    rq_activate_all_grippers(True)
    # end: URCap Program Node
  end
  $ 58 "zero_ftsensor()"
  zero_ftsensor()
  $ 59 "EXTT"
  $ 60 "Set GRP_3F_Enable=Off"
  set_standard_digital_out(4, False)
  $ 61 "Set BarcodeTrigger=Off"
  set_standard_digital_out(6, False)
  $ 62 "Set GRP_3F_Decap=Off"
  set_standard_digital_out(3, False)
  $ 63 "Set GRP_3F_Cap=Off"
  set_standard_digital_out(2, False)
  $ 64 "Set GRP_3F_Open=Off"
  set_standard_digital_out(5, False)
  $ 65 "PSE_T≔get_tool_free_pose(dir=[0,0,0.150], move_in_base_frame=True)"
  global PSE_T=get_tool_free_pose(dir=[0,0,0.150], move_in_base_frame=True)
  $ 66 "If is_reachable(Base_const, [PSE_T])"
  if (is_reachable(p[0.0,0.0,0.0,0.0,0.0,0.0], [PSE_T])):
    $ 67 "MoveL"
    $ 68 "PSE_T" "breakAfter"
    movel(PSE_T, a=1.2, v=0.15)
  end
  $ 69 "powder dispensing variable init"
  $ 70 "Start_thread≔ False "
  global Start_thread=  False
  $ 71 "vib_thread≔ False "
  global vib_thread=  False
  $ 72 "w_full_thread≔ False "
  global w_full_thread=  False
  $ 73 "Picking≔ False "
  global Picking=  False
  $ 74 "d_cc≔0.07"
  global d_cc=0.07
  $ 75 "kp≔0.0035"
  global kp=0.0035
  $ 76 "ki≔0.0001"
  global ki=0.0001
  $ 77 "kd≔0.003"
  global kd=0.003
  $ 78 "dt≔0.2"
  global dt=0.2
  $ 79 "Integral_error≔0"
  global Integral_error=0
  $ 80 "current_error≔0"
  global current_error=0
  $ 81 "previous_error≔0"
  global previous_error=0
  $ 82 "tilt_increment≔0"
  global tilt_increment=0
  $ 83 "tilt_angle≔0"
  global tilt_angle=0
  $ 84 "diff≔0"
  global diff=0
  $ 85 "tilt_to_home()"
  tilt_to_home()
  $ 86 "params_init()"
  params_init()
  $ 87 "switch_spat_M≔ True "
  global switch_spat_M=  True
  $ 88 "switch_spat_S≔ True "
  global switch_spat_S=  True
  $ 89 "switch_spat_F_M≔ True "
  global switch_spat_F_M=  True
  $ 90 "switch_spat_F_S≔ True "
  global switch_spat_F_S=  True
  $ 861 "Thread_1"
  thread Thread_1():
    while (True):
      $ 862 "Dosing Weight"
      $ 863 "If Start_thread≟ True "
      if (Start_thread ==   True  ):
        $ 864 "weight_value≔get_weight()"
        global weight_value=get_weight()
        $ 865 "diff≔target_weight-weight_value"
        global diff=target_weight-weight_value
        $ 866 "Wait: 0.2"
        sleep(0.2)
        $ 867 "sync()"
        sync()
      end
      $ 868 "sync()"
      sync()
    end
  end
  threadId_Thread_1 = run Thread_1()
  $ 869 "Thread_2"
  thread Thread_2():
    while (True):
      $ 883 "Vibration motor"
      $ 884 "Loop vib_thread≟ True "
      thread Thread_while_884():
        while (True):
          $ 885 "If spatula≟'spatula_S' "
          global thread_flag_885=0
          thread Thread_if_885():
            $ 886 "vibration_4()"
            vibration_4()
            thread_flag_885 = 1
          end
          if (spatula == "spatula_S" ):
            global thread_handler_885=run Thread_if_885()
            while (thread_flag_885 == 0):
              if not(spatula == "spatula_S" ):
                kill thread_handler_885
                thread_flag_885 = 2
              else:
                sync()
              end
            end
          else:
            thread_flag_885 = 2
          end
          if (thread_flag_885 == 2):
            $ 887 "ElseIf spatula≟'spatula_M'"
            if (spatula == "spatula_M"):
              $ 888 "vibration_3()"
              vibration_3()
            else:
              $ 889 "Else" "noBreak"
              $ 890 "Set AO[0]=0.0"
              set_standard_analog_out(0, 0.0)
              $ 891 "textmsg('stopped')"
              textmsg("stopped")
            end
          end
        end
      end
      if (vib_thread ==   True  ):
        global thread_handler_884=run Thread_while_884()
        while (vib_thread ==   True  ):
          sync()
        end
        kill thread_handler_884
      end
      $ 892 "sync()"
      sync()
    end
  end
  threadId_Thread_2 = run Thread_2()
  $ 893 "Thread_3"
  thread Thread_3():
    while (True):
      $ 894 "Container weight"
      $ 895 "If w_full_thread≟ True "
      if (w_full_thread ==   True  ):
        $ 896 "aa_weight_cont≔get_cont_weight()"
        global aa_weight_cont=get_cont_weight()
        $ 897 "Wait: 0.2"
        sleep(0.2)
        $ 898 "sync()"
        sync()
      end
      $ 899 "sync()"
      sync()
    end
  end
  threadId_Thread_3 = run Thread_3()
  while (True):
    $ 92 "Robot Program"
    $ 93 "MAIN"
    $ 94 "command_manager(external_control='uGO', cond_suspend=(ITM_Manipulated and AMR_AtTarget and AMR_Charging and AMR_Battery<40), cond_unsuspend=(AMR_Battery≟60))"
    command_manager(external_control="uGO", cond_suspend=(ITM_Manipulated  and  AMR_AtTarget  and  AMR_Charging  and  AMR_Battery<40), cond_unsuspend=(AMR_Battery == 60))
    $ 95 "log_state(STATE_Info)"
    log_state(STATE_Info)
    $ 96 "Switch STATE"
    switch_1 = STATE
    $ 97 "Case 1"
    if (1 == switch_1):
      $ 98 "Stopping"
      $ 99 "STATE_Info≔'Stopping'"
      global STATE_Info="Stopping"
      $ 100 "end_freedrive_mode()"
      end_freedrive_mode()
      $ 101 "Set"
      set_tcp(p[0.0,0.0,0.161,3.1415,0.0,0.0])
      $ 102 "PSE_T≔get_tool_free_pose(dir=[0,0,0.150], move_in_base_frame=True)"
      global PSE_T=get_tool_free_pose(dir=[0,0,0.150], move_in_base_frame=True)
      $ 103 "If is_reachable(Base_const, [PSE_T])"
      if (is_reachable(p[0.0,0.0,0.0,0.0,0.0,0.0], [PSE_T])):
        $ 104 "MoveL"
        $ 105 "PSE_T" "breakAfter"
        movel(PSE_T, a=1.2, v=0.15)
      end
      $ 106 "do_transition(keep_rxry=OBJ_Picked, r=0)"
      do_transition(keep_rxry=OBJ_Picked, r=0)
      $ 115 "Call Sub_AMR_MiR_V3"
      Sub_AMR_MiR_V3()
      $ 116 "If stopping() and AMR_Done"
      if (stopping()  and  AMR_Done):
        $ 117 "STATE≔2"
        global STATE=2
        $ 118 "ugo_update_outputs()"
        ugo_update_outputs()
      end
    elif (2 == switch_1):
      $ 119 "Case 2"
      $ 120 "Stopped"
      $ 121 "STATE_Info≔'Stopped'"
      global STATE_Info="Stopped"
      $ 122 "Call Sub_AMR_MiR_V3"
      Sub_AMR_MiR_V3()
      $ 123 "If CMD_Reset  or PB_Start"
      if (CMD_Reset   or  get_standard_digital_in(0)):
        $ 124 "STATE≔3"
        global STATE=3
        $ 125 "ugo_update_outputs()"
        ugo_update_outputs()
      end
    elif (3 == switch_1):
      $ 126 "Case 3"
      $ 127 " Resetting"
      $ 128 "STATE_Info≔'Resetting'"
      global STATE_Info="Resetting"
      $ 129 "uML"
      $ 130 "reset_error()"
      reset_error()
      $ 131 "reset_warning()"
      reset_warning()
      $ 132 "PROCESS_Step≔0"
      global PROCESS_Step=0
      $ 133 "PROCESS_Info≔''"
      global PROCESS_Info=""
      $ 134 "ARM_Referenced≔ False "
      global ARM_Referenced=  False
      $ 135 "WRK_Done≔ False "
      global WRK_Done=  False
      $ 136 "ITM_Prepared≔ False "
      global ITM_Prepared=  False
      $ 137 "ITM_Manipulated≔ False "
      global ITM_Manipulated=  False
      $ 138 "STP≔0"
      global STP=0
      $ 139 "Action≔0"
      global Action=0
      $ 140 "Action_Info≔''"
      global Action_Info=""
      $ 141 "ITM_ID≔0"
      global ITM_ID=0
      $ 142 "JIG≔0"
      global JIG=0
      $ 143 "JIG_Slot≔0"
      global JIG_Slot=0
      $ 144 "Task_info≔''"
      global Task_info=""
      $ 145 "Set"
      set_tcp(p[0.0,0.0,0.161,3.1415,0.0,0.0])
      $ 146 "App"
      $ 147 "'ADD APPLICATION SPECIFIC COMMANDS'"
      # 'ADD APPLICATION SPECIFIC COMMANDS'
      $ 148 "OBJ_Type≔0"
      global OBJ_Type=0
      $ 149 "OBJ_Nbr≔0"
      global OBJ_Nbr=0
      $ 150 "If CNT_Rack_Output≥50"
      if (CNT_Rack_Output >= 50):
        $ 151 "CNT_Rack_Output≔0"
        global CNT_Rack_Output=0
      end
      $ 152 "TASK≔struct(ID=0, NAVI=struct(target=0, footprint=0, protectiveOff=0, dock=0), WORK=struct(ITM_ID_Src=0, JIG_ID_Src=0, OBJ_Nbr_Src=0, ACT_Src=0, ITM_ID_Tgt=0, JIG_ID_Tgt=0, OBJ_Nbr_Tgt=0, ACT_Tgt=0, OBJ_Type=0))"
      global TASK=struct(ID=0, NAVI=struct(target=0, footprint=0, protectiveOff=0, dock=0), WORK=struct(ITM_ID_Src=0, JIG_ID_Src=0, OBJ_Nbr_Src=0, ACT_Src=0, ITM_ID_Tgt=0, JIG_ID_Tgt=0, OBJ_Nbr_Tgt=0, ACT_Tgt=0, OBJ_Type=0))
      $ 153 "Call Sub_AMR_MiR_V3"
      Sub_AMR_MiR_V3()
      $ 154 "If resetting() and AMR_Done"
      if (resetting()  and  AMR_Done):
        $ 155 "STATE≔4"
        global STATE=4
        $ 156 "ugo_update_outputs()"
        ugo_update_outputs()
      end
    elif (4 == switch_1):
      $ 157 "Case 4"
      $ 158 "Idle"
      $ 159 "STATE_Info≔'Idle'"
      global STATE_Info="Idle"
      $ 160 "If CMD_Start"
      if (CMD_Start):
        $ 161 "STATE≔5"
        global STATE=5
        $ 162 "ugo_update_outputs()"
        ugo_update_outputs()
      end
    elif (5 == switch_1):
      $ 163 "Case 5"
      $ 164 "Starting"
      $ 165 "STATE_Info≔'Starting'"
      global STATE_Info="Starting"
      $ 166 "'ADD COMMANDS WHAT TO START WITH'"
      # 'ADD COMMANDS WHAT TO START WITH'
      $ 167 "Call Sub_AMR_MiR_V3"
      Sub_AMR_MiR_V3()
      $ 168 "get ugo data"
      $ 169 "Assign Tasks"
      $ 170 "TASK.ID = ugo_get_task()"
      TASK.ID = ugo_get_task()
      $ 171 "If TASK.ID≟1"
      if (TASK.ID == 1):
        $ 172 "Task_info≔'Charge'"
        global Task_info="Charge"
        $ 173 "Parameters"
        $ 174 "AMR_PosTarget≔1"
        global AMR_PosTarget=1
      else:
        $ 175 "ElseIf TASK.ID≟9"
        if (TASK.ID == 9):
          $ 176 "'Pick Sarstedt Rack from Variable source'"
          # 'Pick Sarstedt Rack from Variable source'
          $ 177 "Task_info≔'Navigate to Target'"
          global Task_info="Navigate to Target"
          $ 178 "Parameters"
          $ 179 "AMR_PosTarget≔UGO.read_input('00','ITM_ID')"
          global AMR_PosTarget=UGO.read_input("00","ITM_ID")
        else:
          $ 180 "ElseIf TASK.ID≟13"
          if (TASK.ID == 13):
            $ 181 "Task_info≔'Dose Powder'"
            global Task_info="Dose Powder"
            $ 182 "Parameters"
            $ 183 "ITM_ID≔1"
            global ITM_ID=1
            $ 184 "W_now≔(UGO.read_input('00','Container_weight'))/1000"
            global W_now=(UGO.read_input("00","Container_weight"))/1000
            $ 185 "Pow_name≔(UGO.read_input('00','Powder_name'))"
            global Pow_name=(UGO.read_input("00","Powder_name"))
            $ 186 "target_weight≔(UGO.read_input('00','Target_weight'))/1000"
            global target_weight=(UGO.read_input("00","Target_weight"))/1000
            $ 187 "params_init()"
            params_init()
            $ 188 "send_picking_info(Pow_name,target_weight)"
            send_picking_info(Pow_name,target_weight)
            $ 190 "OBJ_Type≔6"
            global OBJ_Type=6
            $ 191 "JIG≔17"
            global JIG=17
            $ 192 "AMR_PosTarget≔5"
            global AMR_PosTarget=5
          else:
            $ 193 "ElseIf TASK.ID≟49"
            if (TASK.ID == 49):
              $ 194 "Task_info≔'Pick Containers'"
              global Task_info="Pick Containers"
              $ 195 "Parameters"
              $ 196 "ITM_ID≔1"
              global ITM_ID=1
              $ 197 "OBJ_Type≔6"
              global OBJ_Type=6
              $ 198 "JIG≔15"
              global JIG=15
              $ 199 "AMR_PosTarget≔3"
              global AMR_PosTarget=3
            else:
              $ 200 "ElseIf TASK.ID≟50"
              if (TASK.ID == 50):
                $ 201 "Task_info≔'Decap Containers'"
                global Task_info="Decap Containers"
                $ 202 "Parameters"
                $ 203 "ITM_ID≔1"
                global ITM_ID=1
                $ 204 "OBJ_Type≔6"
                global OBJ_Type=6
                $ 205 "JIG≔16"
                global JIG=16
                $ 206 "AMR_PosTarget≔5"
                global AMR_PosTarget=5
              else:
                $ 207 "ElseIf TASK.ID≟51"
                if (TASK.ID == 51):
                  $ 208 "Task_info≔'Detect Spatula and transfer powder'"
                  global Task_info="Detect Spatula and transfer powder"
                  $ 209 "Parameters"
                  $ 210 "ITM_ID≔1"
                  global ITM_ID=1
                  $ 211 "target_weight≔(UGO.read_input('00','Target_weight'))/1000"
                  global target_weight=(UGO.read_input("00","Target_weight"))/1000
                  $ 212 "OBJ_Type≔8"
                  global OBJ_Type=8
                  $ 213 "JIG≔16"
                  global JIG=16
                  $ 214 "AMR_PosTarget≔5"
                  global AMR_PosTarget=5
                else:
                  $ 215 "ElseIf TASK.ID≟52"
                  if (TASK.ID == 52):
                    $ 216 "Task_info≔'Pick Powder'"
                    global Task_info="Pick Powder"
                    $ 217 "Parameters"
                    $ 218 "ITM_ID≔1"
                    global ITM_ID=1
                    $ 220 "OBJ_Type≔6"
                    global OBJ_Type=6
                    $ 221 "JIG≔15"
                    global JIG=15
                    $ 222 "AMR_PosTarget≔3"
                    global AMR_PosTarget=3
                  else:
                    $ 223 "ElseIf TASK.ID≟53"
                    if (TASK.ID == 53):
                      $ 224 "Task_info≔'Decap Powder'"
                      global Task_info="Decap Powder"
                      $ 225 "Parameters"
                      $ 226 "ITM_ID≔1"
                      global ITM_ID=1
                      $ 227 "OBJ_Type≔6"
                      global OBJ_Type=6
                      $ 228 "JIG≔1"
                      global JIG=1
                      $ 229 "AMR_PosTarget≔5"
                      global AMR_PosTarget=5
                    else:
                      $ 230 "ElseIf TASK.ID≟54"
                      if (TASK.ID == 54):
                        $ 231 "Task_info≔'Empty and swap Powder container'"
                        global Task_info="Empty and swap Powder container"
                        $ 240 "Parameters"
                        $ 241 "ITM_ID≔1"
                        global ITM_ID=1
                        $ 243 "W_now≔(UGO.read_input('00','Container_weight'))/1000"
                        global W_now=(UGO.read_input("00","Container_weight"))/1000
                        $ 244 "Pow_name≔(UGO.read_input('00','Powder_name'))"
                        global Pow_name=(UGO.read_input("00","Powder_name"))
                        $ 247 "OBJ_Type≔6"
                        global OBJ_Type=6
                        $ 248 "JIG≔17"
                        global JIG=17
                        $ 249 "AMR_PosTarget≔5"
                        global AMR_PosTarget=5
                      else:
                        $ 250 "ElseIf TASK.ID≟55"
                        if (TASK.ID == 55):
                          $ 251 "Task_info≔'Place Powder'"
                          global Task_info="Place Powder"
                          $ 252 "Parameters"
                          $ 253 "ITM_ID≔1"
                          global ITM_ID=1
                          $ 254 "OBJ_Type≔6"
                          global OBJ_Type=6
                          $ 255 "JIG≔21"
                          global JIG=21
                          $ 256 "AMR_PosTarget≔5"
                          global AMR_PosTarget=5
                        else:
                          $ 257 "ElseIf TASK.ID≟56"
                          if (TASK.ID == 56):
                            $ 258 "Task_info≔'Dose Powder'"
                            global Task_info="Dose Powder"
                            $ 259 "Parameters"
                            $ 260 "ITM_ID≔1"
                            global ITM_ID=1
                            $ 261 "target_weight≔(UGO.read_input('00','Target_weight'))/1000"
                            global target_weight=(UGO.read_input("00","Target_weight"))/1000
                            $ 262 "W_now≔(UGO.read_input('00','Container_weight'))/1000"
                            global W_now=(UGO.read_input("00","Container_weight"))/1000
                            $ 263 "Pow_name≔(UGO.read_input('00','Powder_name'))"
                            global Pow_name=(UGO.read_input("00","Powder_name"))
                            $ 264 "OBJ_Type≔6"
                            global OBJ_Type=6
                            $ 265 "JIG≔17"
                            global JIG=17
                            $ 266 "AMR_PosTarget≔5"
                            global AMR_PosTarget=5
                          else:
                            $ 267 "ElseIf TASK.ID≟57"
                            if (TASK.ID == 57):
                              $ 268 "Task_info≔'Recipe Powder dosing'"
                              global Task_info="Recipe Powder dosing"
                              $ 269 "Parameters"
                              $ 270 "ITM_ID≔1"
                              global ITM_ID=1
                              $ 271 "Pow_A≔(UGO.read_input('00','PowderA'))"
                              global Pow_A=(UGO.read_input("00","PowderA"))
                              $ 272 "Pow_B≔(UGO.read_input('00','PowderB'))"
                              global Pow_B=(UGO.read_input("00","PowderB"))
                              $ 273 "Pow_C≔(UGO.read_input('00','PowderC'))"
                              global Pow_C=(UGO.read_input("00","PowderC"))
                              $ 274 "Total_weight≔(UGO.read_input('00','Total_weight'))/1000"
                              global Total_weight=(UGO.read_input("00","Total_weight"))/1000
                              $ 275 "Pow_A_percent≔(UGO.read_input('00','PowderA_percentage'))/100"
                              global Pow_A_percent=(UGO.read_input("00","PowderA_percentage"))/100
                              $ 276 "Pow_B_percent≔(UGO.read_input('00','PowderB_percentage'))/100"
                              global Pow_B_percent=(UGO.read_input("00","PowderB_percentage"))/100
                              $ 277 "Pow_C_percent≔(UGO.read_input('00','PowderC_percentage'))/100"
                              global Pow_C_percent=(UGO.read_input("00","PowderC_percentage"))/100
                              $ 278 "OBJ_Type≔6"
                              global OBJ_Type=6
                              $ 279 "JIG≔17"
                              global JIG=17
                              $ 280 "AMR_PosTarget≔5"
                              global AMR_PosTarget=5
                            else:
                              $ 281 "ElseIf TASK.ID≟58"
                              if (TASK.ID == 58):
                                $ 282 "Task_info≔'Pick Powder containers'"
                                global Task_info="Pick Powder containers"
                                $ 283 "Parameters"
                                $ 284 "ITM_ID≔1"
                                global ITM_ID=1
                                $ 285 "OBJ_Type≔6"
                                global OBJ_Type=6
                                $ 286 "JIG≔15"
                                global JIG=15
                                $ 287 "AMR_PosTarget≔3"
                                global AMR_PosTarget=3
                              else:
                                $ 288 "ElseIf TASK.ID≟59"
                                if (TASK.ID == 59):
                                  $ 289 "Task_info≔'Empty Powder container'"
                                  global Task_info="Empty Powder container"
                                  $ 290 "Parameters"
                                  $ 291 "ITM_ID≔1"
                                  global ITM_ID=1
                                  $ 293 "Pow_name≔(UGO.read_input('00','Powder_name'))"
                                  global Pow_name=(UGO.read_input("00","Powder_name"))
                                  $ 295 "target_weight≔(aa_weight_cont-empty_weight_g)"
                                  global target_weight=(aa_weight_cont-empty_weight_g)
                                  $ 296 "W_now≔target_weight"
                                  global W_now=target_weight
                                  $ 297 "params_init()"
                                  params_init()
                                  $ 298 "send_picking_info(Pow_name,target_weight)"
                                  send_picking_info(Pow_name,target_weight)
                                  $ 299 "w_dosed_total≔0"
                                  global w_dosed_total=0
                                  $ 300 "OBJ_Type≔6"
                                  global OBJ_Type=6
                                  $ 301 "JIG≔17"
                                  global JIG=17
                                  $ 302 "AMR_PosTarget≔5"
                                  global AMR_PosTarget=5
                                else:
                                  $ 303 "ElseIf TASK.ID≟61"
                                  if (TASK.ID == 61):
                                    $ 304 "Task_info≔'Weigh, Place & Decap'"
                                    global Task_info="Weigh, Place & Decap"
                                    $ 305 "Parameters"
                                    $ 306 "ITM_ID≔1"
                                    global ITM_ID=1
                                    $ 307 "OBJ_Type≔6"
                                    global OBJ_Type=6
                                    $ 308 "JIG≔21"
                                    global JIG=21
                                    $ 309 "AMR_PosTarget≔5"
                                    global AMR_PosTarget=5
                                  else:
                                    $ 310 "ElseIf TASK.ID≟62"
                                    if (TASK.ID == 62):
                                      $ 311 "Task_info≔'Dose Powder'"
                                      global Task_info="Dose Powder"
                                      $ 312 "Parameters"
                                      $ 313 "ITM_ID≔1"
                                      global ITM_ID=1
                                      $ 315 "W_now≔aa_weight_cont"
                                      global W_now=aa_weight_cont
                                      $ 316 "Pow_name≔(UGO.read_input('00','Powder_name'))"
                                      global Pow_name=(UGO.read_input("00","Powder_name"))
                                      $ 317 "target_weight≔(UGO.read_input('00','Target_weight'))/1000"
                                      global target_weight=(UGO.read_input("00","Target_weight"))/1000
                                      $ 319 "params_init()"
                                      params_init()
                                      $ 320 "send_picking_info(Pow_name,target_weight)"
                                      send_picking_info(Pow_name,target_weight)
                                      $ 321 "OBJ_Type≔6"
                                      global OBJ_Type=6
                                      $ 322 "JIG≔17"
                                      global JIG=17
                                      $ 323 "AMR_PosTarget≔5"
                                      global AMR_PosTarget=5
                                    else:
                                      $ 324 "ElseIf TASK.ID≟64"
                                      if (TASK.ID == 64):
                                        $ 325 "Task_info≔'Dosing Fumehood'"
                                        global Task_info="Dosing Fumehood"
                                        $ 326 "Parameters"
                                        $ 327 "ITM_ID≔1"
                                        global ITM_ID=1
                                        $ 328 "W_now≔(UGO.read_input('00','Container_weight'))/1000"
                                        global W_now=(UGO.read_input("00","Container_weight"))/1000
                                        $ 329 "OBJ_Type≔6"
                                        global OBJ_Type=6
                                        $ 330 "JIG≔21"
                                        global JIG=21
                                        $ 331 "AMR_PosTarget≔6"
                                        global AMR_PosTarget=6
                                      else:
                                        $ 332 "Else" "noBreak"
                                        $ 333 "set_error(ERROR_WRONG_ORDER)"
                                        set_error(ERROR_WRONG_ORDER)
                                      end
                                    end
                                  end
                                end
                              end
                            end
                          end
                        end
                      end
                    end
                  end
                end
              end
            end
          end
        end
      end
      $ 334 "test ugo"
      $ 335 "Wait: 0.2"
      sleep(0.2)
      $ 336 "ugo_update_outputs()"
      ugo_update_outputs()
      $ 337 "If starting() and AMR_Done"
      if (starting()  and  AMR_Done):
        $ 338 "log_message(Task_info, 'New Task: ')"
        log_message(Task_info, "New Task: ")
        $ 339 "log_message(to_str(TASK.ID), 'Task_ID: ')"
        log_message(to_str(TASK.ID), "Task_ID: ")
        $ 340 "do_transition(keep_rxry=OBJ_Picked)"
        do_transition(keep_rxry=OBJ_Picked)
        $ 341 "STATE≔6"
        global STATE=6
        $ 342 "ugo_update_outputs()"
        ugo_update_outputs()
      end
    elif (6 == switch_1):
      $ 343 "Case 6"
      $ 344 "Execute"
      $ 345 "STATE_Info≔'Execute'"
      global STATE_Info="Execute"
      $ 346 "If  not CMD_Hold and not CMD_Suspend"
      global thread_flag_346=0
      thread Thread_if_346():
        $ 347 "Switch PROCESS_Step"
        switch_2 = PROCESS_Step
        $ 348 "Case 0"
        if (0 == switch_2):
          $ 349 "PROCESS_Info≔'process control'"
          global PROCESS_Info="process control"
          $ 350 "log_process(PROCESS_Info)"
          log_process(PROCESS_Info)
          $ 351 "process control"
          $ 352 "If  not AMR_AtTarget"
          if (  not  AMR_AtTarget):
            $ 353 "PROCESS_Step≔1"
            global PROCESS_Step=1
          else:
            $ 354 "ElseIf (( not ITM_Prepared and  not WRK_Done) or (ITM_Prepared and WRK_Done))"
            if (((  not  ITM_Prepared  and    not  WRK_Done)  or  (ITM_Prepared  and  WRK_Done))):
              $ 355 "PROCESS_Step≔2"
              global PROCESS_Step=2
            else:
              $ 356 "ElseIf  not WRK_Done"
              if (  not  WRK_Done):
                $ 357 "PROCESS_Step≔3"
                global PROCESS_Step=3
              else:
                $ 358 "Else" "noBreak"
                $ 359 "task finished"
                $ 360 "PROCESS_Info≔''"
                global PROCESS_Info=""
                $ 361 "STATE≔7"
                global STATE=7
                $ 362 "ugo_update_outputs()"
                ugo_update_outputs()
              end
            end
          end
        elif (1 == switch_2):
          $ 363 "Case 1"
          $ 364 "navigate"
          $ 365 "'MOVING THE uML'"
          # 'MOVING THE uML'
          $ 366 "PROCESS_Info≔'move to target'"
          global PROCESS_Info="move to target"
          $ 367 "log_process(PROCESS_Info)"
          log_process(PROCESS_Info)
          $ 368 "If TASK.ID≟1"
          if (TASK.ID == 1):
            $ 369 "Action≔51"
            global Action=51
          else:
            $ 370 "Else" "noBreak"
            $ 371 "Action≔52"
            global Action=52
          end
          $ 372 "Call Sub_AMR_MiR_V3"
          Sub_AMR_MiR_V3()
          $ 373 "If AMR_Done"
          if (AMR_Done):
            $ 374 "PROCESS_Step≔0"
            global PROCESS_Step=0
          end
        elif (2 == switch_2):
          $ 375 "Case 2"
          $ 376 "prepare"
          $ 377 "'THINGS THAT HAVE TO BE DONE ONCE IN A SEQUENCE,WORKFLOW'"
          # 'THINGS THAT HAVE TO BE DONE ONCE IN A SEQUENCE,WORKFLOW'
          $ 378 "PROCESS_Info≔'prepare for work'"
          global PROCESS_Info="prepare for work"
          $ 379 "log_process(PROCESS_Info)"
          log_process(PROCESS_Info)
          $ 380 "If TASK.WORK.ITM_ID_Src>1"
          if (TASK.WORK.ITM_ID_Src>1):
            $ 381 "ITM_ID≔TASK.WORK.ITM_ID_Src"
            global ITM_ID=TASK.WORK.ITM_ID_Src
          else:
            $ 382 "ElseIf TASK.WORK.ITM_ID_Tgt>1"
            if (TASK.WORK.ITM_ID_Tgt>1):
              $ 383 "ITM_ID≔TASK.WORK.ITM_ID_Tgt"
              global ITM_ID=TASK.WORK.ITM_ID_Tgt
            end
          end
          $ 384 "If  not ARM_Referenced and (ITM_ID≠0)"
          if (  not  ARM_Referenced  and  (ITM_ID != 0)):
            $ 385 "STP≔1"
            global STP=1
          else:
            $ 386 "ElseIf ARM_Referenced or (ITM_ID≟0)"
            if (ARM_Referenced  or  (ITM_ID == 0)):
              $ 387 "STP≔2"
              global STP=2
            end
          end
          $ 388 "Switch STP"
          switch_3 = STP
          $ 389 "Case 1"
          if (1 == switch_3):
            $ 390 "reference"
            $ 391 "STP_Info≔'reference at target position'"
            global STP_Info="reference at target position"
            $ 392 "log_step(STP_Info)"
            log_step(STP_Info)
            $ 393 "If ITM_ID≟1"
            if (ITM_ID == 1):
              $ 394 "CAM_Done≔ True "
              global CAM_Done=  True
            else:
              $ 395 "Else" "noBreak"
              $ 396 "Action≔131"
              global Action=131
              $ 397 "Call Sub_Vision_V18"
              Sub_Vision_V18()
            end
            $ 399 "If CAM_Done and  not ERROR.FLAG"
            if (CAM_Done  and    not  ERROR.FLAG):
              $ 400 "log_step('ARM referenced')"
              log_step("ARM referenced")
              $ 401 "ARM_Referenced≔ True "
              global ARM_Referenced=  True
            end
          elif (2 == switch_3):
            $ 402 "Case 2"
            $ 403 "manipulate"
            $ 404 "STP_Info≔'manipulate item'"
            global STP_Info="manipulate item"
            $ 405 "log_step(STP_Info)"
            log_step(STP_Info)
            $ 406 "'In case pressing button is needed'"
            # 'In case pressing button is needed'
            $ 407 "If found_in_list(ITM_ID, ITM_ID_List)"
            if (found_in_list(ITM_ID, ITM_ID_List)):
              $ 408 "Switch ITM_ID"
              switch_4 = ITM_ID
              $ 409 "Case 0"
              if (0 == switch_4):
                $ 410 "ITM_Manipulated≔ not ITM_Manipulated"
                global ITM_Manipulated=  not  ITM_Manipulated
              elif (1 == switch_4):
                $ 411 "Case 1"
                $ 412 "ITM_Manipulated≔ not ITM_Manipulated"
                global ITM_Manipulated=  not  ITM_Manipulated
              elif (2 == switch_4):
                $ 413 "Case 2"
              else:
                $ 423 "Default Case"
                $ 424 "ITM_Manipulated≔ not ITM_Manipulated"
                global ITM_Manipulated=  not  ITM_Manipulated
              end
            end
          end
          $ 425 "ITM_Prepared≔(ITM_Manipulated or  not found_in_list(ITM_ID, ITM_ID_List)) and (ARM_Referenced or ITM_ID≟0) and  not WRK_Done"
          global ITM_Prepared=(ITM_Manipulated  or    not  found_in_list(ITM_ID, ITM_ID_List))  and  (ARM_Referenced  or  ITM_ID == 0)  and    not  WRK_Done
          $ 426 "STP≔0"
          global STP=0
          $ 427 "STP_Info≔''"
          global STP_Info=""
          $ 428 "PROCESS_Step≔0"
          global PROCESS_Step=0
        elif (3 == switch_2):
          $ 429 "Case 3"
          $ 430 "work"
          $ 431 "'ADD EVERY MACHINE, OBJECT, STATION TO WORK ON'"
          # 'ADD EVERY MACHINE, OBJECT, STATION TO WORK ON'
          $ 432 "Switch ITM_ID"
          switch_3 = ITM_ID
          $ 433 "Case 1"
          if (1 == switch_3):
            $ 434 "uLM"
            $ 435 "If TASK.ID≟12"
            if (TASK.ID == 12):
              $ 436 "fill racks"
              $ 437 "Action≔151"
              global Action=151
              $ 438 "Call Sub_Vision_V18"
              Sub_Vision_V18()
              $ 439 "If  not ERROR.FLAG"
              if (  not  ERROR.FLAG):
                $ 440 "Actions for the task"
                $ 441 "Action≔1"
                global Action=1
                $ 442 "JIG≔2"
                global JIG=2
                $ 443 "JIG_Slot≔CAM_Result[0]"
                global JIG_Slot=CAM_Result[0]
                $ 444 "OBJ_Nbr≔CAM_Result[0]"
                global OBJ_Nbr=CAM_Result[0]
                $ 445 "OBJ_Type≔2"
                global OBJ_Type=2
                $ 446 "Call Sub_Action_V4"
                Sub_Action_V4()
                $ 447 "If OBJ_Picked"
                if (OBJ_Picked):
                  $ 448 "CAM_Result.remove(0)"
                  CAM_Result.remove(0)
                  $ 449 "PRC_TubCounter≔PRC_TubCounter+1"
                  global PRC_TubCounter=PRC_TubCounter+1
                  $ 450 "If PRC_TubCounter%4≟0"
                  if (PRC_TubCounter%4 == 0):
                    $ 451 "JIG_Slot≔4"
                    global JIG_Slot=4
                  else:
                    $ 452 "Else" "noBreak"
                    $ 453 "JIG_Slot≔PRC_TubCounter%4"
                    global JIG_Slot=PRC_TubCounter%4
                  end
                  $ 454 "OBJ_Nbr≔ceil(PRC_TubCounter/4)"
                  global OBJ_Nbr=ceil(PRC_TubCounter/4)
                  $ 455 "Action≔2"
                  global Action=2
                  $ 456 "JIG≔4"
                  global JIG=4
                  $ 457 "Call Sub_Action_V4"
                  Sub_Action_V4()
                  $ 458 "Action≔151"
                  global Action=151
                  $ 459 "Call Sub_Vision_V18"
                  Sub_Vision_V18()
                end
              end
              $ 460 "If (CAM_Captures≥CAM_PRM_Retries) or (PRC_TubCounter≥32)"
              if ((CAM_Captures >= CAM_PRM_Retries)  or  (PRC_TubCounter >= 32)):
                $ 461 "PROCESS_Step≔0"
                global PROCESS_Step=0
                $ 462 "WRK_Done≔ True "
                global WRK_Done=  True
              end
            else:
              $ 463 "ElseIf TASK.ID≟13"
              if (TASK.ID == 13):
                $ 464 "Dose Powder"
                $ 465 "Action≔131"
                global Action=131
                $ 466 "Call Sub_Vision_V18"
                Sub_Vision_V18()
                $ 467 "Action≔34"
                global Action=34
                $ 468 "Call Sub_Action_V4"
                Sub_Action_V4()
                $ 469 "PROCESS_Step≔0"
                global PROCESS_Step=0
                $ 470 "WRK_Done≔ True "
                global WRK_Done=  True
              else:
                $ 471 "ElseIf TASK.ID≟49"
                if (TASK.ID == 49):
                  $ 472 "Pick Powder container"
                  $ 473 "Action≔131"
                  global Action=131
                  $ 474 "Call Sub_Vision_V18"
                  Sub_Vision_V18()
                  $ 475 "Action≔35"
                  global Action=35
                  $ 476 "Call Sub_Action_V4"
                  Sub_Action_V4()
                  $ 477 "PROCESS_Step≔0"
                  global PROCESS_Step=0
                  $ 478 "WRK_Done≔ True "
                  global WRK_Done=  True
                else:
                  $ 479 "ElseIf TASK.ID≟50"
                  if (TASK.ID == 50):
                    $ 480 "Decap containers"
                    $ 481 "Action≔36"
                    global Action=36
                    $ 482 "Call Sub_Action_V4"
                    Sub_Action_V4()
                    $ 483 "PROCESS_Step≔0"
                    global PROCESS_Step=0
                    $ 484 "WRK_Done≔ True "
                    global WRK_Done=  True
                  else:
                    $ 485 "ElseIf TASK.ID≟51"
                    if (TASK.ID == 51):
                      $ 486 "Detect Spatula and transfer powder"
                      $ 487 "Action≔131"
                      global Action=131
                      $ 488 "Call Sub_Vision_V18"
                      Sub_Vision_V18()
                      $ 489 "Action≔37"
                      global Action=37
                      $ 490 "Call Sub_Action_V4"
                      Sub_Action_V4()
                      $ 491 "PROCESS_Step≔0"
                      global PROCESS_Step=0
                      $ 492 "WRK_Done≔ True "
                      global WRK_Done=  True
                    else:
                      $ 493 "ElseIf TASK.ID≟52"
                      if (TASK.ID == 52):
                        $ 494 "Pick Powder container"
                        $ 495 "Action≔131"
                        global Action=131
                        $ 496 "Call Sub_Vision_V18"
                        Sub_Vision_V18()
                        $ 497 "Action≔39"
                        global Action=39
                        $ 498 "Call Sub_Action_V4"
                        Sub_Action_V4()
                        $ 499 "PROCESS_Step≔0"
                        global PROCESS_Step=0
                        $ 500 "WRK_Done≔ True "
                        global WRK_Done=  True
                      else:
                        $ 501 "ElseIf TASK.ID≟53"
                        if (TASK.ID == 53):
                          $ 502 "Decap containerA"
                          $ 503 "Action≔40"
                          global Action=40
                          $ 504 "Call Sub_Action_V4"
                          Sub_Action_V4()
                          $ 505 "PROCESS_Step≔0"
                          global PROCESS_Step=0
                          $ 506 "WRK_Done≔ True "
                          global WRK_Done=  True
                        else:
                          $ 507 "ElseIf TASK.ID≟55"
                          if (TASK.ID == 55):
                            $ 508 "Place Powder"
                            $ 509 "Action≔131"
                            global Action=131
                            $ 510 "Call Sub_Vision_V18"
                            Sub_Vision_V18()
                            $ 511 "Action≔41"
                            global Action=41
                            $ 512 "Call Sub_Action_V4"
                            Sub_Action_V4()
                            $ 513 "PROCESS_Step≔0"
                            global PROCESS_Step=0
                            $ 514 "WRK_Done≔ True "
                            global WRK_Done=  True
                          else:
                            $ 515 "ElseIf TASK.ID≟54"
                            if (TASK.ID == 54):
                              $ 516 "Empty and swap container"
                              $ 517 "Action≔131"
                              global Action=131
                              $ 518 "Call Sub_Vision_V18"
                              Sub_Vision_V18()
                              $ 519 "Action≔42"
                              global Action=42
                              $ 520 "Call Sub_Action_V4"
                              Sub_Action_V4()
                              $ 521 "PROCESS_Step≔0"
                              global PROCESS_Step=0
                              $ 522 "WRK_Done≔ True "
                              global WRK_Done=  True
                            else:
                              $ 523 "ElseIf TASK.ID≟56"
                              if (TASK.ID == 56):
                                $ 524 "Dispense Powder"
                                $ 525 "Action≔131"
                                global Action=131
                                $ 526 "Call Sub_Vision_V18"
                                Sub_Vision_V18()
                                $ 527 "Action≔43"
                                global Action=43
                                $ 528 "Call Sub_Action_V4"
                                Sub_Action_V4()
                                $ 529 "PROCESS_Step≔0"
                                global PROCESS_Step=0
                                $ 530 "WRK_Done≔ True "
                                global WRK_Done=  True
                              else:
                                $ 531 "ElseIf TASK.ID≟57"
                                if (TASK.ID == 57):
                                  $ 532 "Recipe Dosing"
                                  $ 533 "Action≔48"
                                  global Action=48
                                  $ 534 "Call Sub_Action_V4"
                                  Sub_Action_V4()
                                  $ 551 "PROCESS_Step≔0"
                                  global PROCESS_Step=0
                                  $ 552 "WRK_Done≔ True "
                                  global WRK_Done=  True
                                else:
                                  $ 553 "ElseIf TASK.ID≟58"
                                  if (TASK.ID == 58):
                                    $ 554 "Pick Powder containers"
                                    $ 555 "Num_cont_picked≔0"
                                    global Num_cont_picked=0
                                    $ 556 "powder_position≔'Position1'"
                                    global powder_position="Position1"
                                    $ 557 "Loop Num_cont_picked<3"
                                    while (Num_cont_picked<3):
                                      $ 558 "Action≔131"
                                      global Action=131
                                      $ 559 "Call Sub_Vision_V18"
                                      Sub_Vision_V18()
                                      $ 560 "Action≔47"
                                      global Action=47
                                      $ 561 "Call Sub_Action_V4"
                                      Sub_Action_V4()
                                    end
                                    $ 562 "PROCESS_Step≔0"
                                    global PROCESS_Step=0
                                    $ 563 "WRK_Done≔ True "
                                    global WRK_Done=  True
                                  else:
                                    $ 564 "ElseIf TASK.ID≟59"
                                    if (TASK.ID == 59):
                                      $ 565 "Empty powder container"
                                      $ 566 "Action≔131"
                                      global Action=131
                                      $ 567 "Call Sub_Vision_V18"
                                      Sub_Vision_V18()
                                      $ 568 "Action≔50"
                                      global Action=50
                                      $ 569 "Call Sub_Action_V4"
                                      Sub_Action_V4()
                                      $ 570 "PROCESS_Step≔0"
                                      global PROCESS_Step=0
                                      $ 571 "WRK_Done≔ True "
                                      global WRK_Done=  True
                                    else:
                                      $ 572 "ElseIf TASK.ID≟61"
                                      if (TASK.ID == 61):
                                        $ 573 "Place Powder"
                                        $ 574 "Action≔131"
                                        global Action=131
                                        $ 575 "Call Sub_Vision_V18"
                                        Sub_Vision_V18()
                                        $ 576 "Action≔51"
                                        global Action=51
                                        $ 577 "Call Sub_Action_V4"
                                        Sub_Action_V4()
                                        $ 578 "PROCESS_Step≔0"
                                        global PROCESS_Step=0
                                        $ 579 "WRK_Done≔ True "
                                        global WRK_Done=  True
                                      else:
                                        $ 580 "ElseIf TASK.ID≟62"
                                        if (TASK.ID == 62):
                                          $ 581 "Dose Powder"
                                          $ 582 "Action≔131"
                                          global Action=131
                                          $ 583 "Call Sub_Vision_V18"
                                          Sub_Vision_V18()
                                          $ 584 "Action≔52"
                                          global Action=52
                                          $ 585 "Call Sub_Action_V4"
                                          Sub_Action_V4()
                                          $ 586 "PROCESS_Step≔0"
                                          global PROCESS_Step=0
                                          $ 587 "WRK_Done≔ True "
                                          global WRK_Done=  True
                                        else:
                                          $ 588 "ElseIf TASK.ID≟64"
                                          if (TASK.ID == 64):
                                            $ 589 "Fumehood Powder dose"
                                            $ 590 "Action≔131"
                                            global Action=131
                                            $ 591 "Call Sub_Vision_V18"
                                            Sub_Vision_V18()
                                            $ 592 "Action≔54"
                                            global Action=54
                                            $ 593 "Call Sub_Action_V4"
                                            Sub_Action_V4()
                                            $ 594 "PROCESS_Step≔0"
                                            global PROCESS_Step=0
                                            $ 595 "WRK_Done≔ True "
                                            global WRK_Done=  True
                                          end
                                        end
                                      end
                                    end
                                  end
                                end
                              end
                            end
                          end
                        end
                      end
                    end
                  end
                end
              end
            end
          elif (2 == switch_3):
            $ 596 "Case 2"
          elif (5 == switch_3):
            $ 638 "Case 5"
          elif (20 == switch_3):
            $ 646 "Case 20"
          elif (43 == switch_3):
            $ 708 "Case 43"
          else:
            $ 716 "Default Case"
            $ 717 "WRK_Done≔ True "
            global WRK_Done=  True
            $ 718 "PROCESS_Step≔0"
            global PROCESS_Step=0
          end
        end
        thread_flag_346 = 1
      end
      if (  not  CMD_Hold and not CMD_Suspend):
        global thread_handler_346=run Thread_if_346()
        while (thread_flag_346 == 0):
          if not(  not  CMD_Hold and not CMD_Suspend):
            kill thread_handler_346
            thread_flag_346 = 2
          else:
            sync()
          end
        end
      else:
        thread_flag_346 = 2
      end
      $ 719 "If CMD_Hold"
      if (CMD_Hold):
        $ 720 "STATE≔9"
        global STATE=9
        $ 721 "ugo_update_outputs()"
        ugo_update_outputs()
      else:
        $ 722 "ElseIf CMD_Suspend"
        if (CMD_Suspend):
          $ 723 "STATE≔12"
          global STATE=12
          $ 724 "ugo_update_outputs()"
          ugo_update_outputs()
        end
      end
    elif (7 == switch_1):
      $ 725 "Case 7"
      $ 726 "Completing"
      $ 727 "STATE_Info≔'Completing'"
      global STATE_Info="Completing"
      $ 728 "'ADD COMMANDS FOR COMPLETING THE PROCESS'"
      # 'ADD COMMANDS FOR COMPLETING THE PROCESS'
      $ 729 "do_transition(keep_rxry=OBJ_Picked)"
      do_transition(keep_rxry=OBJ_Picked)
      $ 730 "Call Sub_AMR_MiR_V3"
      Sub_AMR_MiR_V3()
      $ 731 "If completing() and AMR_Done"
      if (completing()  and  AMR_Done):
        $ 732 "STATE≔8"
        global STATE=8
        $ 733 "ugo_update_outputs()"
        ugo_update_outputs()
      end
    elif (8 == switch_1):
      $ 734 "Case 8"
      $ 735 "Complete"
      $ 736 "STATE_Info≔'Complete'"
      global STATE_Info="Complete"
      $ 737 "If CMD_Reset"
      if (CMD_Reset):
        $ 738 "STATE≔3"
        global STATE=3
        $ 739 "ugo_update_outputs()"
        ugo_update_outputs()
      end
    elif (9 == switch_1):
      $ 740 "Case 9"
      $ 741 "Holding"
      $ 742 "STATE_Info≔'Holding'"
      global STATE_Info="Holding"
      $ 743 "stopl(0.5)"
      stopl(0.5)
      $ 744 "Call Sub_AMR_MiR_V3"
      Sub_AMR_MiR_V3()
      $ 745 "If holding() and AMR_Done"
      if (holding()  and  AMR_Done):
        $ 746 "STATE≔10"
        global STATE=10
        $ 747 "ugo_update_outputs()"
        ugo_update_outputs()
      end
    elif (10 == switch_1):
      $ 748 "Case 10"
      $ 749 "Held"
      $ 750 "STATE_Info≔'Held'"
      global STATE_Info="Held"
      $ 751 "If CMD_Unhold"
      if (CMD_Unhold):
        $ 752 "end_freedrive_mode()"
        end_freedrive_mode()
        $ 753 "STATE≔11"
        global STATE=11
        $ 754 "ugo_update_outputs()"
        ugo_update_outputs()
      else:
        $ 755 "ElseIf FNC_Freedrive"
        if (FNC_Freedrive):
          $ 756 "freedrive_mode()"
          freedrive_mode()
        else:
          $ 757 "Else" "noBreak"
          $ 758 "end_freedrive_mode()"
          end_freedrive_mode()
        end
      end
    elif (11 == switch_1):
      $ 759 "Case 11"
      $ 760 "Unholding"
      $ 761 "STATE_Info≔'Unholding'"
      global STATE_Info="Unholding"
      $ 762 "Clearing"
      $ 763 "Switch ERROR.ID"
      switch_2 = ERROR.ID
      $ 764 "Case 1002"
      if (1002 == switch_2):
        $ 765 "AMR_AtTarget≔ False "
        global AMR_AtTarget=  False
        $ 766 "ARM_Referenced≔ False "
        global ARM_Referenced=  False
        $ 767 "ITM_Prepared≔ False "
        global ITM_Prepared=  False
        $ 768 "PROCESS_Step≔1"
        global PROCESS_Step=1
      elif (2007 == switch_2):
        $ 769 "Case 2007"
        $ 770 "PROCESS_Step≔1"
        global PROCESS_Step=1
      end
      $ 771 "reset_error()"
      reset_error()
      $ 772 "reset_warning()"
      reset_warning()
      $ 773 "OBJ_Picked≔gripper_has_object()"
      global OBJ_Picked=gripper_has_object()
      $ 774 "Call Sub_AMR_MiR_V3"
      Sub_AMR_MiR_V3()
      $ 775 "If unholding() and AMR_Done"
      if (unholding()  and  AMR_Done):
        $ 776 "STATE≔6"
        global STATE=6
        $ 777 "ugo_update_outputs()"
        ugo_update_outputs()
      end
    elif (12 == switch_1):
      $ 778 "Case 12"
      $ 779 "Suspending"
      $ 780 "STATE_Info≔'Suspending'"
      global STATE_Info="Suspending"
      $ 781 "PROCESS_Info≔str_cat(PROCESS_Info, ' suspended')"
      global PROCESS_Info=str_cat(PROCESS_Info, " suspended")
      $ 782 "If suspending()"
      if (suspending()):
        $ 783 "STATE≔13"
        global STATE=13
        $ 784 "ugo_update_outputs()"
        ugo_update_outputs()
      end
    elif (13 == switch_1):
      $ 785 "Case 13"
      $ 786 "Suspended"
      $ 787 "STATE_Info≔'Suspended'"
      global STATE_Info="Suspended"
      $ 788 "Call Sub_AMR_MiR_V3"
      Sub_AMR_MiR_V3()
      $ 789 "If CMD_Unsuspend"
      if (CMD_Unsuspend):
        $ 790 "STATE≔14"
        global STATE=14
        $ 791 "ugo_update_outputs()"
        ugo_update_outputs()
      end
    elif (14 == switch_1):
      $ 792 "Case 14"
      $ 793 "Unsuspending"
      $ 794 "STATE_Info≔'Unsuspending'"
      global STATE_Info="Unsuspending"
      $ 795 "PROCESS_Step≔0"
      global PROCESS_Step=0
      $ 796 "If unsuspending()"
      if (unsuspending()):
        $ 797 "STATE≔6"
        global STATE=6
        $ 798 "ugo_update_outputs()"
        ugo_update_outputs()
      end
    elif (15 == switch_1):
      $ 799 "Case 15"
      $ 800 "Aborting"
      $ 801 "STATE_Info≔'Aborting'"
      global STATE_Info="Aborting"
      $ 802 "If aborting()"
      if (aborting()):
        $ 803 "STATE≔16"
        global STATE=16
        $ 804 "ugo_update_outputs()"
        ugo_update_outputs()
      end
    elif (16 == switch_1):
      $ 805 "Case 16"
      $ 806 "Aborted"
      $ 807 "STATE_Info≔'Aborted'"
      global STATE_Info="Aborted"
      $ 808 "If CMD_Clear"
      if (CMD_Clear):
        $ 809 "STATE≔17"
        global STATE=17
        $ 810 "ugo_update_outputs()"
        ugo_update_outputs()
      end
    elif (17 == switch_1):
      $ 811 "Case 17"
      $ 812 "Clearing"
      $ 813 "STATE_Info≔'Clearing'"
      global STATE_Info="Clearing"
      $ 814 "Clearing"
      $ 815 "reset_warning()"
      reset_warning()
      $ 816 "reset_error()"
      reset_error()
      $ 817 "If clearing()"
      if (clearing()):
        $ 818 "STATE≔2"
        global STATE=2
        $ 819 "ugo_update_outputs()"
        ugo_update_outputs()
      end
    end
    $ 820 "log_state(STATE_Info)"
    log_state(STATE_Info)
    $ 821 "log_warning(WARNING.MSG)"
    log_warning(WARNING.MSG)
    $ 822 "log_error(ERROR.MSG)"
    log_error(ERROR.MSG)
    $ 823 "Times"
    $ 824 "Switch STATE"
    switch_1 = STATE
    $ 825 "Case 1"
    if (1 == switch_1):
      $ 826 "TM_St_Stopping≔get_time(STATE_Times[STATE-1])"
      global TM_St_Stopping=get_time(STATE_Times[STATE-1])
    elif (2 == switch_1):
      $ 827 "Case 2"
      $ 828 "TM_St_Stopped≔get_time(STATE_Times[STATE-1])"
      global TM_St_Stopped=get_time(STATE_Times[STATE-1])
    elif (3 == switch_1):
      $ 829 "Case 3"
      $ 830 "TM_St_Resetting≔get_time(STATE_Times[STATE-1])"
      global TM_St_Resetting=get_time(STATE_Times[STATE-1])
    elif (4 == switch_1):
      $ 831 "Case 4"
      $ 832 "TM_St_Idle≔get_time(STATE_Times[STATE-1])"
      global TM_St_Idle=get_time(STATE_Times[STATE-1])
    elif (5 == switch_1):
      $ 833 "Case 5"
      $ 834 "TM_St_Starting≔get_time(STATE_Times[STATE-1])"
      global TM_St_Starting=get_time(STATE_Times[STATE-1])
    elif (6 == switch_1):
      $ 835 "Case 6"
      $ 836 "TM_St_Execute≔get_time(STATE_Times[STATE-1])"
      global TM_St_Execute=get_time(STATE_Times[STATE-1])
    elif (7 == switch_1):
      $ 837 "Case 7"
      $ 838 "TM_St_Completin≔get_time(STATE_Times[STATE-1])"
      global TM_St_Completin=get_time(STATE_Times[STATE-1])
    elif (8 == switch_1):
      $ 839 "Case 8"
      $ 840 "TM_St_Complete≔get_time(STATE_Times[STATE-1])"
      global TM_St_Complete=get_time(STATE_Times[STATE-1])
    elif (9 == switch_1):
      $ 841 "Case 9"
      $ 842 "TM_St_Holding≔get_time(STATE_Times[STATE-1])"
      global TM_St_Holding=get_time(STATE_Times[STATE-1])
    elif (10 == switch_1):
      $ 843 "Case 10"
      $ 844 "TM_St_Held≔get_time(STATE_Times[STATE-1])"
      global TM_St_Held=get_time(STATE_Times[STATE-1])
    elif (11 == switch_1):
      $ 845 "Case 11"
      $ 846 "TM_St_Unholding≔get_time(STATE_Times[STATE-1])"
      global TM_St_Unholding=get_time(STATE_Times[STATE-1])
    elif (12 == switch_1):
      $ 847 "Case 12"
      $ 848 "TM_St_Suspendin≔get_time(STATE_Times[STATE-1])"
      global TM_St_Suspendin=get_time(STATE_Times[STATE-1])
    elif (13 == switch_1):
      $ 849 "Case 13"
      $ 850 "TM_St_Suspended≔get_time(STATE_Times[STATE-1])"
      global TM_St_Suspended=get_time(STATE_Times[STATE-1])
    elif (14 == switch_1):
      $ 851 "Case 14"
      $ 852 "TM_St_Unsuspend≔get_time(STATE_Times[STATE-1])"
      global TM_St_Unsuspend=get_time(STATE_Times[STATE-1])
    elif (15 == switch_1):
      $ 853 "Case 15"
      $ 854 "TM_St_Aborting≔get_time(STATE_Times[STATE-1])"
      global TM_St_Aborting=get_time(STATE_Times[STATE-1])
    elif (16 == switch_1):
      $ 855 "Case 16"
      $ 856 "TM_St_Aborted≔get_time(STATE_Times[STATE-1])"
      global TM_St_Aborted=get_time(STATE_Times[STATE-1])
    elif (17 == switch_1):
      $ 857 "Case 17"
      $ 858 "TM_St_Clearing≔get_time(STATE_Times[STATE-1])"
      global TM_St_Clearing=get_time(STATE_Times[STATE-1])
    end
    $ 860 "Wait: 0.1"
    sleep(0.1)
  end
end
